SUBAPPLICATION Uebung_OPC_L10_AX (* Wie Training_10, lokal: Input_I1/I2 (Hoch/Runter) per lokalem PUBLISH, ILOCK schaltet Output_Q7/Q8 *)
  (* Standard: 61499-2; Description: Copyright (c) 2026 Meisterschulen am Ostbahnhof This program and the accompanying materials are made available under the terms of the Eclipse Public License 2.0 which is available at https://www.eclipse.org/legal/epl-2.0/ SPDX-License-Identifier: EPL-2.0 *)
  (* Version 1.0, 2026-10-18, Franz Höpfinger, Meisterschulen am Ostbahnhof, Aus SubApp_PC_A + SubApp_PC_B von test_VV zusammengefuehrt, lokale Varianten der Bausteine *)
  PACKAGE Meins::OPC_UA_Lokal;
  IMPORT Meins::OPC_UA_Lokal::const::OpcUaLokal::SW1_UP_WRITE;
  IMPORT Meins::OPC_UA_Lokal::const::OpcUaLokal::SW1_DOWN_WRITE;
  IMPORT logiBUS::io::DI::logiBUS_DI::Input_I1;
  IMPORT logiBUS::io::DI::logiBUS_DI::Input_I2;
  IMPORT Meins::OPC_UA_Lokal::const::OpcUaLokal::SW1_UP_READ;
  IMPORT Meins::OPC_UA_Lokal::const::OpcUaLokal::SW1_DOWN_READ;
  IMPORT logiBUS::io::DQ::logiBUS_DO::Output_Q7;
  IMPORT logiBUS::io::DQ::logiBUS_DO::Output_Q8;
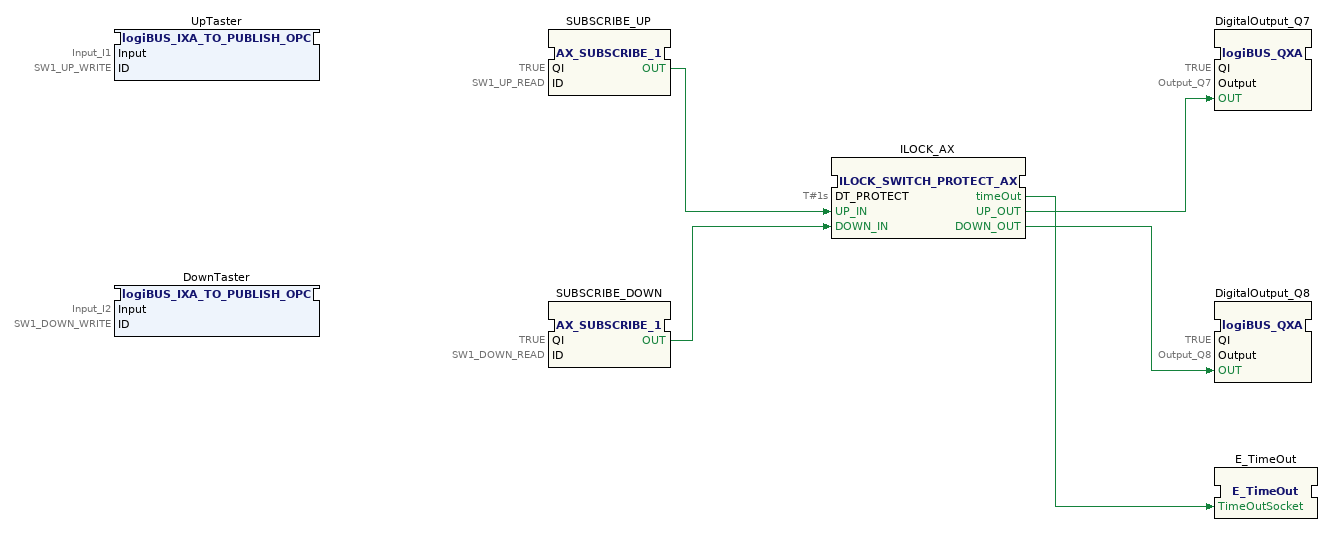
  FBS
    SUBSCRIBE_UP : adapter::net::AX_SUBSCRIBE_1(QI := TRUE, ID := SW1_UP_READ);
    SUBSCRIBE_DOWN : adapter::net::AX_SUBSCRIBE_1(QI := TRUE, ID := SW1_DOWN_READ);
    ILOCK_AX : logiBUS::signalprocessing::interlock::ILOCK_SWITCH_PROTECT_AX(DT_PROTECT := T#1s);
    E_TimeOut : iec61499::events::E_TimeOut;
    DigitalOutput_Q7 : logiBUS::io::DQ::logiBUS_QXA(QI := TRUE, Output := Output_Q7);
    DigitalOutput_Q8 : logiBUS::io::DQ::logiBUS_QXA(QI := TRUE, Output := Output_Q8);
  END_FBS
  SUBAPPS
    UpTaster : MyLib::sys::logiBUS_IXA_TO_PUBLISH_OPC(Input := Input_I1, ID := SW1_UP_WRITE);
    DownTaster : MyLib::sys::logiBUS_IXA_TO_PUBLISH_OPC(Input := Input_I2, ID := SW1_DOWN_WRITE);
  END_SUBAPPS
  ADAPTER_CONNECTIONS
    SUBSCRIBE_UP.OUT TO ILOCK_AX.UP_IN;
    SUBSCRIBE_DOWN.OUT TO ILOCK_AX.DOWN_IN;
    ILOCK_AX.timeOut TO E_TimeOut.TimeOutSocket;
    ILOCK_AX.UP_OUT TO DigitalOutput_Q7.OUT;
    ILOCK_AX.DOWN_OUT TO DigitalOutput_Q8.OUT;
  END_CONNECTIONS
END_SUBAPPLICATION
